(* IEC 61131-3 sources: plc-vscode/tests/st/all/rusty/tests/lit/single/pointer, 33 files *)

(* ---- reference_to_array_of_pointers_assignment.st ---- *)
// RUN: (%COMPILE %s && %RUN) | %CHECK %s
TYPE userType :
    DINT := 0;
END_TYPE

FUNCTION main : DINT
    VAR
        x : userType := 101;
        y : userType := 202;
        z : userType := 303;
        w : userType := 404;

        a : REFERENCE TO ARRAY [1..2] OF POINTER TO userType;
        b : ARRAY [1..2] OF POINTER TO userType;
        c : ARRAY [1..2] OF POINTER TO userType;
        d : ARRAY [1..2] OF POINTER TO userType;
    END_VAR

    // b starts as z/w, d starts as x/y
    b[1] := ADR(z);
    b[2] := ADR(w);
    c[1] := ADR(z);
    c[2] := ADR(w);
    d[1] := ADR(x);
    d[2] := ADR(y);

    // 1) REF= binds reference to target array variable (a -> d)
    a REF= d;

    // 2) b := a reads through reference and copies dereferenced array value
    b := a;

    // CHECK: b-after-b:=a 101 202
    printf('b-after-b:=a %d %d$N', b[1]^, b[2]^);

    // 3) a := c writes into referenced array (d := c)
    a := c;

    // CHECK: d-after-a:=c 303 404
    printf('d-after-a:=c %d %d$N', d[1]^, d[2]^);

    // Keep exact bug-report statements as compile-time/runtime no-op checks
    a REF= b;
    b := a;
    a := b;

    // CHECK: after-bug-sequence 101 202
    printf('after-bug-sequence %d %d$N', b[1]^, b[2]^);
END_FUNCTION

(* ---- referenceto_variable_referencing_struct.st ---- *)
// RUN: (%COMPILE %s && %RUN) | %CHECK %s
TYPE Transaction : STRUCT
    id      : DINT;
    amount  : DINT;
    message : STRING;
END_STRUCT END_TYPE

FUNCTION main : DINT
    VAR
        txn     : Transaction := (id := 1, amount := 5, message := 'whats up');
        refTxn  : REFERENCE TO Transaction;
    END_VAR

    refTxn REF= txn;

    // CHECK: 1
    printf('%d$N', refTxn.id);

    // CHECK: 5
    printf('%d$N', refTxn.amount);

    // CHECK: whats up
    printf('%s$N', REF(refTxn.message));
END_FUNCTION

(* ---- paren_ref_arith_deref.st ---- *)
// RUN: (%COMPILE %s && %RUN) | %CHECK %s
// Regression for #1443: pointer arithmetic on a paren-REF result followed by
// a deref must read the adjacent slot, not segfault.

FUNCTION main : DINT
VAR
    arr : ARRAY[0..1] OF DINT := [10, 20];
    out_val : DINT;
END_VAR
    out_val := (REF(arr[0]) + 1)^;
    // CHECK: 20
    printf('%d$N', out_val);
    main := 0;
END_FUNCTION

(* ---- paren_ref_deref_assign.st ---- *)
// RUN: (%COMPILE %s && %RUN) | %CHECK %s
// Regression for #1463: writing through `(REF(x))^ := value` must reach `x`
// instead of segfaulting. The codegen change extracts the pointer directly
// from the RValue produced by REF instead of loading through it.

FUNCTION main : DINT
VAR
    x : DINT := 0;
END_VAR
    (REF(x))^ := 99;
    // CHECK: 99
    printf('%d$N', x);
    main := 0;
END_FUNCTION

(* ---- paren_ref_deref_read.st ---- *)
// RUN: (%COMPILE %s && %RUN) | %CHECK %s
// Regression for #1443: reading through `(REF(x))^` must dereference the
// returned pointer, not load through the variable holding it. Prior to the
// fix this silently miscompiled to a segfault at runtime.

FUNCTION main : DINT
VAR
    x : DINT := 42;
    y : DINT;
END_VAR
    y := (REF(x))^;
    // CHECK: 42
    printf('%d$N', y);
    main := 0;
END_FUNCTION

(* ---- pointer_to_return_not_affected_by_ref_lowering.st ---- *)
// RUN: (%COMPILE %s && %RUN) | %CHECK %s
// Regression test: ensure reference-to-return lowering does not affect POINTER TO returns.
// A function returning POINTER TO INT should keep its return type and continue to work
// normally rather than being lowered as though it returned REFERENCE TO.
FUNCTION getPointer : POINTER TO INT
    VAR_INPUT
        in	: REF_TO INT;
    END_VAR

    getPointer := in;
END_FUNCTION

FUNCTION main : DINT
    VAR
        ptr    : POINTER TO INT;
        tmpVal : INT := 42;
    END_VAR

    ptr := getPointer(REF(tmpVal));

    // CHECK: 42
    printf('%d$N', ptr^);
END_FUNCTION

(* ---- ref_assignment_operator.st ---- *)
// RUN: (%COMPILE %s && %RUN) | %CHECK %s
FUNCTION main : DINT
    VAR
        a : REF_TO DINT;
        b : DINT := 5;
    END_VAR
    a REF= b;

    // CHECK: 5
    printf('%d$N', a^);
END_FUNCTION

(* ---- ref_assignment_with_parenthesis.st ---- *)
// RUN: (%COMPILE %s && %RUN) | %CHECK %s
FUNCTION main : DINT
    VAR
        refe: REFERENCE TO DINT;
        myDint : DINT;
    END_VAR

    myDint := 10;
    refe REF= (myDint);

    // CHECK: 10
    printf('%d$N', refe);
END_FUNCTION

(* ---- ref_to_return_not_affected_by_ref_lowering.st ---- *)
// RUN: (%COMPILE %s && %RUN) | %CHECK %s
// Regression test: functions returning REF_TO must not be rewritten by the
// reference-to-return lowering.
FUNCTION getRef : REF_TO INT
    VAR_INPUT
        in	: REF_TO INT;
    END_VAR

    getRef := in;
END_FUNCTION

FUNCTION main : DINT
    VAR
        ptr    : REF_TO INT;
        tmpVal : INT := 77;
    END_VAR

    ptr := getRef(REF(tmpVal));

    // CHECK: 77
    printf('%d$N', ptr^);
END_FUNCTION

(* ---- reference_to_null.st ---- *)
// RUN: (%COMPILE %s && %RUN) | %CHECK %s
FUNCTION main: DINT
    VAR
        foo : REFERENCE TO DINT;
        foo2 : REFERENCE TO INT;
        bar,baz,qux : DINT;
    END_VAR

    // Set to null
    foo REF= 0;
    // Should not crash

    // Set to null
    foo2 REF= 0;
    // Should not crash

    foo REF= bar;
    bar := 1;
    baz := 2;
    qux := 2;

    // CHECK: 2
    bar := bar + foo; // bar + bar => 1 + 1
    printf('%d$N', foo);

    // CHECK: 4
    baz := baz + foo; // baz + foo => baz + bar => 2 + 2
    foo REF= baz;
    printf('%d$N', foo);

    // CHECK: 6
    qux := qux + foo; // qux + foo => qux + baz => 2 + 4
    foo REF= qux;
    printf('%d$N', foo);

END_FUNCTION

(* ---- referenceto_function_of_type_referenceto.st ---- *)
// RUN: (%COMPILE %s && %RUN) | %CHECK %s
FUNCTION referenceFunc : REFERENCE TO INT
    VAR_INPUT
        in	: REFERENCE TO INT;
    END_VAR

    in := in + 1;
    referenceFunc REF= in;
END_FUNCTION

FUNCTION main : DINT
    VAR
        refVal : REFERENCE TO INT;
        conVal : INT;
        tmpVal : INT;
    END_VAR

    tmpVal := 11;
    refVal REF= tmpVal;
    refVal REF= referenceFunc(refVal);
    conVal := refVal;

    // CHECK: 12
    printf('%d$N', conVal);
END_FUNCTION

(* ---- referenceto_function_of_type_referenceto_aggregate_type.st ---- *)
// RUN: (%COMPILE %s && %RUN) | %CHECK %s
FUNCTION referenceFunc : REFERENCE TO STRING
    VAR_INPUT
        in	: REFERENCE TO STRING;
    END_VAR

    referenceFunc REF= in;
END_FUNCTION

FUNCTION main : DINT
    VAR
        refVal : REFERENCE TO STRING;
        conVal : STRING;
        tmpVal : STRING := 'Hello world!';
    END_VAR

    refVal REF= tmpVal;
    refVal REF= referenceFunc(refVal);
    conVal := refVal;

    // CHECK: Hello world!
    printf('%s$N', conVal);
END_FUNCTION

(* ---- referenceto_function_of_type_referenceto_array.st ---- *)
// RUN: (%COMPILE %s && %RUN) | %CHECK %s
FUNCTION referenceFunc : REFERENCE TO ARRAY[1..3] OF INT
    VAR_INPUT
        in	: REFERENCE TO ARRAY[1..3] OF INT;
    END_VAR

    referenceFunc REF= in;
END_FUNCTION

FUNCTION main : DINT
    VAR
        refVal : REFERENCE TO ARRAY[1..3] OF INT;
        conVal : ARRAY[1..3] OF INT;
        tmpVal : ARRAY[1..3] OF INT;
    END_VAR

    refVal REF= tmpVal;
    tmpVal[1] := 3;
    tmpVal[2] := 2;
    tmpVal[3] := 1;

    refVal REF= referenceFunc(refVal);
    conVal := refVal;

    // CHECK: 1, 2, 3
    printf('%d, %d, %d$N', conVal[3], conVal[2], conVal[1]);
END_FUNCTION

(* ---- referenceto_function_of_type_referenceto_lowered.st ---- *)
// RUN: (%COMPILE %s && %RUN) | %CHECK %s

// Non-lowered code
/*
FUNCTION referenceFunc : REFERENCE TO INT
    VAR_INPUT
        in	: REFERENCE TO INT;
    END_VAR

    in := in + 1;
    referenceFunc REF= in;
END_FUNCTION

FUNCTION main : DINT
    VAR
        refVal : REFERENCE TO INT;
        conVal : INT;
        tmpVal : INT;
    END_VAR

    tmpVal := 11;
    refVal REF= tmpVal;
    refVal REF= referenceFunc(refVal);
    conVal := refVal;
END_FUNCTION
*/

FUNCTION referenceFunc
    VAR_INPUT
        __referenceFunc_return_val : REFERENCE TO INT;
        in	: REFERENCE TO INT;
    END_VAR

    in := in + 1;
    __referenceFunc_return_val := in;
END_FUNCTION

FUNCTION main : DINT
    VAR
        refVal : REFERENCE TO INT;
        conVal : INT;
        tmpVal : INT;
    END_VAR

    VAR_TEMP
        __referenceFunc_return_val : REFERENCE TO INT;
        __referenceFunc_return_val_store : INT;
    END_VAR

    tmpVal := 11;
    refVal REF= tmpVal;
    __referenceFunc_return_val REF= __referenceFunc_return_val_store;
    referenceFunc(__referenceFunc_return_val, refVal);
    refVal REF= __referenceFunc_return_val;
    conVal := refVal;

    // CHECK: 12
    printf('%d$N', conVal);
END_FUNCTION

(* ---- referenceto_return_called_twice.st ---- *)
// RUN: (%COMPILE %s && %RUN) | %CHECK %s
// Verify: calling the same reference-to-return function multiple times at top level.
// The temp variable is shared across calls — verify values don't leak between calls.
FUNCTION referenceFunc : REFERENCE TO INT
    VAR_INPUT
        in	: REFERENCE TO INT;
    END_VAR

    in := in + 1;
    referenceFunc REF= in;
END_FUNCTION

FUNCTION main : DINT
    VAR
        refA   : REFERENCE TO INT;
        refB   : REFERENCE TO INT;
        valA   : INT;
        valB   : INT;
        tmpA   : INT;
        tmpB   : INT;
    END_VAR

    tmpA := 10;
    tmpB := 20;
    refA REF= tmpA;
    refB REF= tmpB;

    refA REF= referenceFunc(refA);  // 10 + 1 = 11
    refB REF= referenceFunc(refB);  // 20 + 1 = 21

    valA := refA;
    valB := refB;

    // CHECK: 11
    printf('%d$N', valA);
    // CHECK: 21
    printf('%d$N', valB);
END_FUNCTION

(* ---- referenceto_return_double_nested_call.st ---- *)
// RUN: (%COMPILE %s && %RUN) | %CHECK %s
// Verify: nested call - result of one ref-return function passed directly to another.
FUNCTION addOne : REFERENCE TO INT
    VAR_INPUT
        in	: REFERENCE TO INT;
    END_VAR

    in := in + 1;
    addOne REF= in;
END_FUNCTION

FUNCTION doubleIt : REFERENCE TO INT
    VAR_INPUT
        in	: REFERENCE TO INT;
    END_VAR

    in := in * 2;
    doubleIt REF= in;
END_FUNCTION

FUNCTION tripleIt : REFERENCE TO INT
    VAR_INPUT
        in	: REFERENCE TO INT;
    END_VAR

    in := in * 3;
    tripleIt REF= in;
END_FUNCTION

FUNCTION main : DINT
    VAR
        refVal : REFERENCE TO INT;
        conVal : INT;
        tmpVal : INT;
    END_VAR

    tmpVal := 5;
    refVal REF= tmpVal;

    // Nested: tripleIt(doubleIt(addOne(refVal))) should give ((5+1)*2)*3 = 36
    refVal REF= tripleIt(doubleIt(addOne(refVal)));
    conVal := refVal;

    // CHECK: 36
    printf('%d$N', conVal);
END_FUNCTION

(* ---- referenceto_return_inside_case.st ---- *)
// RUN: (%COMPILE %s && %RUN) | %CHECK %s
// Test case #2: verify calls inside CASE branches are lowered correctly.
FUNCTION referenceFunc : REFERENCE TO INT
    VAR_INPUT
        in	: REFERENCE TO INT;
    END_VAR

    in := in + 1;
    referenceFunc REF= in;
END_FUNCTION

FUNCTION main : DINT
    VAR
        refVal : REFERENCE TO INT;
        conVal : INT;
        tmpVal : INT;
        sel    : INT := 1;
    END_VAR

    tmpVal := 10;
    refVal REF= tmpVal;

    CASE sel OF
        1:
            refVal REF= referenceFunc(refVal);
        2:
            tmpVal := 99;
    END_CASE;

    conVal := refVal;

    // CHECK: 11
    printf('%d$N', conVal);
END_FUNCTION

(* ---- referenceto_return_inside_for_loop.st ---- *)
// RUN: (%COMPILE %s && %RUN) | %CHECK %s
// Regression test: calls inside FOR loops are lowered correctly.
FUNCTION referenceFunc : REFERENCE TO INT
    VAR_INPUT
        in	: REFERENCE TO INT;
    END_VAR

    in := in + 1;
    referenceFunc REF= in;
END_FUNCTION

FUNCTION main : DINT
    VAR
        refVal : REFERENCE TO INT;
        conVal : INT;
        tmpVal : INT;
        i      : INT;
    END_VAR

    tmpVal := 0;
    refVal REF= tmpVal;

    FOR i := 1 TO 5 DO
        refVal REF= referenceFunc(refVal);
    END_FOR;

    conVal := refVal;

    // CHECK: 5
    printf('%d$N', conVal);
END_FUNCTION

(* ---- referenceto_return_inside_if.st ---- *)
// RUN: (%COMPILE %s && %RUN) | %CHECK %s
// Regression test for critical issue #2: ensure call-site lowering works
// for reference-to-return function calls inside IF control flow.
FUNCTION referenceFunc : REFERENCE TO INT
    VAR_INPUT
        in	: REFERENCE TO INT;
    END_VAR

    in := in + 1;
    referenceFunc REF= in;
END_FUNCTION

FUNCTION main : DINT
    VAR
        refVal : REFERENCE TO INT;
        conVal : INT;
        tmpVal : INT;
        flag   : BOOL := TRUE;
    END_VAR

    tmpVal := 11;
    refVal REF= tmpVal;

    IF flag THEN
        refVal REF= referenceFunc(refVal);
    END_IF;

    conVal := refVal;

    // CHECK: 12
    printf('%d$N', conVal);
END_FUNCTION

(* ---- referenceto_return_inside_while_loop.st ---- *)
// RUN: (%COMPILE %s && %RUN) | %CHECK %s
// Verify calls inside WHILE loops are lowered.
FUNCTION referenceFunc : REFERENCE TO INT
    VAR_INPUT
        in	: REFERENCE TO INT;
    END_VAR

    in := in + 1;
    referenceFunc REF= in;
END_FUNCTION

FUNCTION main : DINT
    VAR
        refVal : REFERENCE TO INT;
        conVal : INT;
        tmpVal : INT;
    END_VAR

    tmpVal := 0;
    refVal REF= tmpVal;

    WHILE refVal < 3 DO
        refVal REF= referenceFunc(refVal);
    END_WHILE;

    conVal := refVal;

    // CHECK: 3
    printf('%d$N', conVal);
END_FUNCTION

(* ---- referenceto_return_multiple_different_functions.st ---- *)
// RUN: (%COMPILE %s && %RUN) | %CHECK %s
// Verify: calling multiple different reference-to-return functions from the same POU.
FUNCTION addOne : REFERENCE TO INT
    VAR_INPUT
        in	: REFERENCE TO INT;
    END_VAR

    in := in + 1;
    addOne REF= in;
END_FUNCTION

FUNCTION doubleIt : REFERENCE TO INT
    VAR_INPUT
        in	: REFERENCE TO INT;
    END_VAR

    in := in * 2;
    doubleIt REF= in;
END_FUNCTION

FUNCTION main : DINT
    VAR
        refVal : REFERENCE TO INT;
        conVal : INT;
        tmpVal : INT;
    END_VAR

    tmpVal := 5;
    refVal REF= tmpVal;

    refVal REF= addOne(refVal);    // 5 + 1 = 6
    refVal REF= doubleIt(refVal);  // 6 * 2 = 12
    conVal := refVal;

    // CHECK: 12
    printf('%d$N', conVal);
END_FUNCTION

(* ---- referenceto_return_nested_call.st ---- *)
// RUN: (%COMPILE %s && %RUN) | %CHECK %s
// Verify: nested call - result of one ref-return function passed directly to another.
FUNCTION addOne : REFERENCE TO INT
    VAR_INPUT
        in	: REFERENCE TO INT;
    END_VAR

    in := in + 1;
    addOne REF= in;
END_FUNCTION

FUNCTION doubleIt : REFERENCE TO INT
    VAR_INPUT
        in	: REFERENCE TO INT;
    END_VAR

    in := in * 2;
    doubleIt REF= in;
END_FUNCTION

FUNCTION main : DINT
    VAR
        refVal : REFERENCE TO INT;
        conVal : INT;
        tmpVal : INT;
    END_VAR

    tmpVal := 5;
    refVal REF= tmpVal;

    // Nested: doubleIt(addOne(refVal)) should give (5+1)*2 = 12
    refVal REF= doubleIt(addOne(refVal));
    conVal := refVal;

    // CHECK: 12
    printf('%d$N', conVal);
END_FUNCTION

(* ---- referenceto_return_not_last_statement.st ---- *)
// RUN: (%COMPILE %s && %RUN) | %CHECK %s
// Regression test for critical issue #3: return lowering must still occur even
// when the REF= assignment to the function name is not the last statement in
// the function body.
FUNCTION referenceFunc : REFERENCE TO INT
    VAR_INPUT
        in	: REFERENCE TO INT;
    END_VAR
    VAR
        dummy : INT;
    END_VAR

    in := in + 1;
    referenceFunc REF= in;
    dummy := 0; // keep a trailing statement to verify the REF= above is still lowered
END_FUNCTION

FUNCTION main : DINT
    VAR
        refVal : REFERENCE TO INT;
        conVal : INT;
        tmpVal : INT;
    END_VAR

    tmpVal := 11;
    refVal REF= tmpVal;
    refVal REF= referenceFunc(refVal);
    conVal := refVal;

    // CHECK: 12
    printf('%d$N', conVal);
END_FUNCTION

(* ---- referenceto_return_standalone_call.st ---- *)
// RUN: (%COMPILE %s && %RUN) | %CHECK %s
// Verify: Standalone calls (without REF= assignment) to reference-to-return
// functions have their signatures rewritten so the call compiles.
// Top-level standalone calls are already handled by this rewriting.
FUNCTION referenceFunc : REFERENCE TO INT
    VAR_INPUT
        in	: REFERENCE TO INT;
    END_VAR

    in := in + 1;
    referenceFunc REF= in;
END_FUNCTION

FUNCTION main : DINT
    VAR
        refVal : REFERENCE TO INT;
        conVal : INT;
        tmpVal : INT;
    END_VAR

    tmpVal := 11;
    refVal REF= tmpVal;

    // Call without capturing the return - should still compile & run with the
    // rewritten void signature (the side effect on `in` still matters)
    referenceFunc(refVal);

    conVal := refVal;

    // CHECK: 12
    printf('%d$N', conVal);
END_FUNCTION

(* ---- referenceto_return_with_early_return.st ---- *)
// RUN: (%COMPILE %s && %RUN) | %CHECK %s
// Regression test: multiple return paths with an early RETURN must preserve
// the REF= assignment to the function name when it occurs in a conditional branch.
FUNCTION selectRef : REFERENCE TO INT
    VAR_INPUT
        a   : REFERENCE TO INT;
        b   : REFERENCE TO INT;
        sel : BOOL;
    END_VAR

    IF sel THEN
        selectRef REF= a;
        RETURN;
    END_IF;

    selectRef REF= b;
END_FUNCTION

FUNCTION main : DINT
    VAR
        refVal : REFERENCE TO INT;
        valA   : INT := 10;
        valB   : INT := 20;
        conVal : INT;
    END_VAR

    refVal REF= valA;

    // sel=TRUE should return reference to valA
    refVal REF= selectRef(refVal, refVal, TRUE);
    conVal := refVal;

    // CHECK: 10
    printf('%d$N', conVal);
END_FUNCTION

(* ---- referenceto_variable_autoderef.st ---- *)
// RUN: (%COMPILE %s && %RUN) | %CHECK %s
FUNCTION main: DINT
    VAR
        foo : REFERENCE TO DINT;
        bar : DINT;
        baz : DINT;
        qux : DINT;
    END_VAR

    foo REF= bar;
    bar := 1;
    baz := 2;
    qux := 2;

    // CHECK: 2
    bar := bar + foo; // bar + bar => 1 + 1
    printf('%d$N', foo);

    // CHECK: 4
    baz := baz + foo; // baz + foo => baz + bar => 2 + 2
    foo REF= baz;
    printf('%d$N', foo);

    // CHECK: 6
    qux := qux + foo; // qux + foo => qux + baz => 2 + 4
    foo REF= qux;
    printf('%d$N', foo);
END_FUNCTION

(* ---- referenceto_variable_referencing_array.st ---- *)
// RUN: (%COMPILE %s && %RUN) | %CHECK %s
FUNCTION main: DINT
    VAR
        arr     :               ARRAY[1..3] OF DINT;
        refArr  : REFERENCE TO  ARRAY[1..3] OF DINT;
    END_VAR

    refArr REF= arr;
    arr[1] := 3;
    arr[2] := 2;
    arr[3] := 1;

    // CHECK: 1, 2, 3
    printf('%d, %d, %d$N', refArr[3], refArr[2], refArr[1]);
END_FUNCTION

(* ---- referenceto_variable_referencing_itself.st ---- *)
// RUN: (%COMPILE %s && %RUN) | %CHECK %s
FUNCTION main : DINT
    VAR
        foo : REFERENCE TO DINT;
        bar : REFERENCE TO DINT;
        qux : DINT;
    END_VAR

    foo REF= bar;
    bar REF= qux;

    bar REF= bar;
    qux := 5;

    // CHECK: 5
    printf('%d$N', bar); // bar (-> bar) -> qux
END_FUNCTION

(* ---- referenceto_variable_referencing_other_referenceto_variable.st ---- *)
// RUN: (%COMPILE %s && %RUN) | %CHECK %s
FUNCTION main : DINT
    VAR
        foo : REFERENCE TO DINT;
        bar : REFERENCE TO DINT;
        qux : DINT;
    END_VAR

    bar REF= qux;
    foo REF= bar;
    qux := 5;

    // CHECK: 5
    printf('%d$N', foo); // foo -> bar -> qux
END_FUNCTION

(* ---- method_call_deref_assign.st ---- *)
// RUN: (%COMPILE %s && %RUN) | %CHECK %s
// Regression for #1463: `methodCall()^ := value` must parse and write through
// the returned pointer. Prior to the fix, the parser closed the call and
// rejected `^` with E007.

FUNCTION_BLOCK Holder
VAR
    x : DINT := 0;
END_VAR
METHOD GetPtr : REF_TO DINT
    GetPtr := REF(x);
END_METHOD
METHOD Read : DINT
    Read := x;
END_METHOD
END_FUNCTION_BLOCK

FUNCTION main : DINT
VAR
    h : Holder;
END_VAR
    h.GetPtr()^ := 17;
    // CHECK: 17
    printf('%d$N', h.Read());
    main := 0;
END_FUNCTION

(* ---- referenceto_return_with_colliding_methods.st ---- *)
// RUN: (%COMPILE %s && %RUN) | %CHECK %s
PROGRAM test
    VAR
        fbIntContainer : fbIntContainer;
        fbIntContainer_value_store : REFERENCE TO IntContainer;
        fbIntContainer_struct_store : IntContainer;

        fbStringContainer : fbStringContainer;
        fbStringContainer_value_store : REFERENCE TO StringContainer;
        fbStringContainer_struct_store : StringContainer;
    END_VAR

    fbIntContainer_struct_store.child := 51;
    fbIntContainer_value_store REF= fbIntContainer_struct_store;
    fbIntContainer.value := fbIntContainer_value_store;

    // CHECK: FB1-Value: 51
    printf('FB1-Value: %d$N', fbIntContainer.value.child);

    fbStringContainer_struct_store.child := 'Hello There';
    fbStringContainer_value_store REF= fbStringContainer_struct_store;
    fbStringContainer.value := fbStringContainer_value_store;

    // CHECK: FB2-Value: Hello There
    printf('FB2-Value: %s$N', fbStringContainer.value.child);
END_PROGRAM

// INT Container
FUNCTION_BLOCK fbIntContainer
    VAR
        _value	: IntContainer;
    END_VAR

    PROPERTY_GET value : REFERENCE TO IntContainer
        value REF= _value;
    END_PROPERTY

    PROPERTY_SET value : REFERENCE TO IntContainer
        _value := value;
    END_PROPERTY
END_FUNCTION_BLOCK

// String Container
FUNCTION_BLOCK fbStringContainer
    VAR
        _value	: StringContainer;
    END_VAR

    PROPERTY_GET value : REFERENCE TO StringContainer
        value REF= _value;
    END_PROPERTY

    PROPERTY_SET value : REFERENCE TO StringContainer
        _value := value;
    END_PROPERTY
END_FUNCTION_BLOCK

TYPE IntContainer :
	STRUCT
		child : INT := 42;
	END_STRUCT
END_TYPE

TYPE StringContainer :
	STRUCT
		child : STRING[255] := 'Hello World';
	END_STRUCT
END_TYPE

FUNCTION main
    test();
END_FUNCTION

(* ---- value_behind_function_block_pointer_is_assigned_to_correctly.st ---- *)
// RUN: (%COMPILE %s && %RUN) | %CHECK %s

FUNCTION_BLOCK file_t
    VAR_INPUT
        var1: BOOL;
        var2: BOOL;
    END_VAR

    VAR_OUTPUT
        out1: BOOL;
        out2: BOOL;
    END_VAR

    out1 := var1;
    out2 := var2;
END_FUNCTION_BLOCK

FUNCTION main: DINT
    VAR
        a: BOOL;
        b: BOOL;
        file: file_t;
        FileOpen: REF_TO file_t;
    END_VAR

    FileOpen := REF(file);
    FileOpen^(var1 := FALSE, var2 := TRUE, out1 => a, out2 => b);

    // CHECK: a = 0
    // CHECK: b = 1
    printf('a = %d$N', a);
    printf('b = %d$N', b);
END_FUNCTION

(* ---- referenceto_struct_resolution_of_types.st ---- *)
// RUN: (%COMPILE %s && %RUN) | %CHECK %s
PROGRAM test
VAR
	myStruct : REFERENCE TO structuredTypeOrFb;
    myStruct_store : structuredTypeOrFb;
END_VAR

myStruct REF= myStruct_store;
printf('%d$N', myStruct.x);

END_PROGRAM

TYPE structuredTypeOrFb :
	STRUCT
		x	: INT := 42;
	END_STRUCT
END_TYPE

FUNCTION main
    // CHECK: 42
    test();
END_FUNCTION
